(*
SPDX-License-Identifier: MIT
License: https://opensource.org/license/mit
*)

(*!
<summary>Runs an owned external element with explicit abort recovery.</summary>
<description>
Owns persistent root instances and fixed child storage. Use from one task without reentry.
Children borrows the same array for the instance lifetime. Root parents remain zero.
</description>
*)

{attribute 'no_assign'}
{attribute 'no_explicit_call' := 'do not call this function block directly'}
FUNCTION_BLOCK ExternalRecoveryTestRunner EXTENDS TOF_Testing.TestRunner<1>
VAR_STAT
	//! <summary>Class name shared by instances of this concrete runner.</summary>
	{attribute 'hide'}
	_ClassName : STRING := __POUNAME();
END_VAR
VAR
	{attribute 'hide'}
	{attribute 'init_namespace'}
	_NamespaceName : STRING;
END_VAR
VAR_OUTPUT
	//! <summary>Owned root element used by this runner.</summary>
	ExternalCase : ExternalElementProbe(name := "External element", parent := 0);
END_VAR
VAR
	_Children : ARRAY [0.._ChildCount - 1] OF TOF_Testing.ITestElement :=
	[
		ExternalCase
	];
END_VAR

(*!
<summary>Borrows the concrete class name; callers must not modify the returned storage.</summary>
*)
{attribute 'monitoring' := 'call'}
PROPERTY ClassName : REFERENCE TO STRING
GET
ClassName REF= _ClassName;
END_GET
END_PROPERTY

(*!
<summary>Borrows the concrete namespace name for the instance lifetime; callers must not modify it.</summary>
*)
{attribute 'monitoring' := 'call'}
PROPERTY NamespaceName : REFERENCE TO STRING
GET
NamespaceName REF= _NamespaceName;
END_GET
END_PROPERTY

(*!
<summary>Reports the complete concrete instance size.</summary>
*)
{attribute 'monitoring' := 'call'}
PROPERTY SelfSize : ULINT
GET
SelfSize := XSIZEOF(THIS^);
END_GET
END_PROPERTY

(*!
<summary>Borrows the unchanged persistent root array; application code must not modify it.</summary>
*)
{attribute 'monitoring' := 'call'}
PROPERTY Children : REFERENCE TO ARRAY [0.._ChildCount - 1] OF TOF_Testing.ITestElement
GET
Children REF= _Children;
END_GET
END_PROPERTY

END_FUNCTION_BLOCK

(* stored: Version 1.1.0.1
   POU ExternalRecoveryTestRunner: Id {a9cf2dc7-84f8-4a82-bf8b-0fcfbc6eb66f}, SpecialFunc None
   Property ClassName: Id {495a5aa3-df4a-4de4-bfeb-a496d70f6f35}
   Get Get: Id {7c31b686-aa0a-4441-b446-67f7094e32c9}
   Property NamespaceName: Id {b74f4f63-11a6-4ae6-a2a7-492ac3c6f9d9}
   Get Get: Id {6ce10ae1-0898-4db8-a581-917279a69dac}
   Property SelfSize: Id {52e9ce12-337d-4b40-9030-33a9e7bc4130}
   Get Get: Id {a4a9e3fa-9422-4b31-b855-1ba5e5b0f6d4}
   Property Children: Id {6c7c508c-70d4-4d74-804e-d9710b0bce74}
   Get Get: Id {33556f14-5c4e-4a06-acfd-238afa8261c8} *)
